Fanuc KAREL source: kt00928.compact.KL

PROGRAM KT00928
%STACKSIZE=65535
%PRIORITY=65535
%NOLOCKGROUP
VAR
S1 : STRING[80]
S2 : STRING[80]
OUT : INTEGER
BEGIN
S1='A'
S2='B'
S1='A'
S2='B'
OUT=ORD(S1,1)
END KT00928
